(* IEC 61131-3 sources: Lasal-MCP/examples/SampleSource/LASALScreenAdvancedSolution/LASALScreenAdvancedSolution/LASALScreenAdvacnedSolution/Stations/Terminal/HMI/Class/MyKeyboardCode, 1 file *)

(* ---- MyKeyboardCode.st ---- *)
(*!
<Class
	Name               = "MyKeyboardCode"
	Revision           = "0.0"
	RealtimeTask       = "false"
	CyclicTask         = "false"
	BackgroundTask     = "false"
	Sigmatek           = "false"
	OSInterface        = "false"
	HighPriority       = "false"
	Automatic          = "false"
	UpdateMode         = "Prescan"
	SharedCommandTable = "true"
	Objectsize         = "(390,180)">
	<Channels>
		<Server Name="KeyCode" Visualized="true" Initialize="false" WriteProtected="true" Retentive="false"/>
	</Channels>
	<Network Name="MyKeyboardCode">
		<!-- List of Components in this network -->
		<Components>
			<Object
				Name       = "_base"
				Class      = "_Global"
				Position   = "(218,120)"
				Visualized = "true"
				Remotely   = "true">
				<Channels>
					<Server Name="Server0"/>
					<Client Name="Lse"/>
				</Channels>
			</Object>
		</Components>
		<Comments>
		</Comments>
		<!-- List of Connections in this network -->
		<Connections>
			<Connection Source="this.Server0" Destination="_base.Server0" Vertices="(690,210),(518,210),"/>
			<Connection Source="_base.Lse" Destination="this.Lse" Vertices="(218,210),(38,210),"/>
		</Connections>
		<!-- Headerfiles -->
		<Options>
		</Options>
	</Network>
</Class>
*)
#pragma using _Global

MyKeyboardCode : CLASS
: _Global
  //Servers:
	KeyCode 	: SvrCh_DINT;
  //Clients:
  //Variables:
  //Functions:

	FUNCTION VIRTUAL GLOBAL IF_WindowRun
		VAR_INPUT
			whoami 	: ^_WHOAMI;
			pic 	: ^void;
			event 	: ^_EVENT;
		END_VAR;
  //Tables:
	FUNCTION @STD
		VAR_OUTPUT
			ret_code	: CONFSTATES;
		END_VAR;
	FUNCTION GLOBAL TAB @CT_;
END_CLASS;

FUNCTION VIRTUAL GLOBAL MyKeyboardCode::IF_WindowRun
	VAR_INPUT
		whoami 	: ^_WHOAMI;
		pic 	: ^void;
		event 	: ^_EVENT;
	END_VAR

  if ((whoami^.ima = IMA_PICTURE) | (whoami^.ima = IMA_WINDOW)) then

    if (event^.ftype = _EVENT_KEYPRESS) then

      KeyCode := event^.scancode;

      //=====================================================
      case KeyCode of
        //---------------------------------------------------
        _F1:  // button F1 to open Screen 1
          InsertCmd(x0:= CMD_NEWPICTURE, x1:= 1, x2:= 0);

        //---------------------------------------------------
        _F2: // button F2 to open Screen 2
          InsertCmd(x0:= CMD_NEWPICTURE, x1:= 2, x2:= 0);

        //---------------------------------------------------
        _F3: // button F3
          InsertCmd(x0:= CMD_NEWPICTURE, x1:= 3, x2:= 0);

        //---------------------------------------------------
        _HOME: // left windows button
          InsertCmd(x0:= CMD_NEWPICTURE, x1:= 0, x2:= 0);

        //---------------------------------------------------
        _ESC: // button ESC
          InsertCmd(x0:= CMD_RETURN, x1:= 0, x2:= 0);

      end_case;
      //=====================================================

    end_if;

  end_if;

END_FUNCTION
